(* IEC 61131-3 sources: plc-workbench/experiments/formal_r7/final_recheck/fault_injection_interlocked_start, 2 files *)

(* ---- before.st ---- *)
FUNCTION_BLOCK InterlockedStart
VAR_INPUT
  start : BOOL;
  stop : BOOL;
  permit : BOOL;
END_VAR
VAR_OUTPUT
  running : BOOL;
END_VAR
VAR
  prevStart : BOOL;
  startEdge : BOOL;
END_VAR

(* Edge detection uses previous scan value; block initial prevStart = FALSE *)
startEdge := start AND NOT prevStart;
prevStart := start;

(* Stop / interlock dominate any simultaneous start edge *)
IF stop OR NOT permit THEN
  running := FALSE;
ELSIF startEdge THEN
  running := TRUE;
END_IF;

END_FUNCTION_BLOCK

(* ---- candidate_final.st ---- *)
FUNCTION_BLOCK InterlockedStart
VAR_INPUT
  start : BOOL;
  stop : BOOL;
  permit : BOOL;
END_VAR
VAR_OUTPUT
  running : BOOL;
END_VAR
VAR
  prevStart : BOOL;
  startEdge : BOOL;
END_VAR

(* Edge detection uses previous scan value; block initial prevStart = FALSE *)
startEdge := start AND NOT prevStart;
prevStart := start;

(* Stop / interlock dominate any simultaneous start edge *)
IF stop OR NOT permit THEN
  running := FALSE;
ELSIF startEdge THEN
  running := TRUE;
END_IF;

END_FUNCTION_BLOCK
